(* PLC project TBEN_L5_PLC11.project, CODESYS CODESYS V3.5 SP21 Patch 1 *)
(* stored: creationDateTime 2026-11-07T15:35:08.08506, modificationDateTime 2026-11-07T15:09:07.4034196 *)

// Ghi DWORD big-endian (4 byte) vào buffer
FUNCTION F_IolSetU32BE : BOOL
VAR_INPUT
    pBuf  : POINTER TO BYTE;
    uiOff : UINT;
    dwVal : DWORD;
END_VAR

            IF pBuf = 0 THEN
    F_IolSetU32BE := FALSE;
    RETURN;
END_IF
F_IolSetU16BE(pBuf, uiOff, DWORD_TO_UINT(SHR(dwVal, 16)));
F_IolSetU16BE(pBuf, uiOff + 2, DWORD_TO_UINT(dwVal));
F_IolSetU32BE := TRUE;

          
END_FUNCTION
